// TIA Portal V20 export
// export: Created 2026-10-19T18:02:39.4342809Z, ExportSetting WithDefaults, DisplayName Totally Integrated Automation Portal, DisplayVersion V20 Update 6, DisplayName TIA Portal Openness, DisplayVersion V20 Update 6, DisplayName TIA Portal Version Control Interface, DisplayVersion V20 Update 6, DisplayName SINAMICS Startdrive Advanced, DisplayVersion V20 SP1, DisplayName SINAMICS Startdrive G130, G150, S120, S150, SINAMICS MV, G220, S200, S210, DisplayVersion V20 SP1, DisplayName SINAMICS Startdrive G110M, G120, G120C, G120D, G120P, G115D, DisplayVersion V20 SP1, DisplayName STEP 7 Professional, DisplayVersion V20 Update 6, DisplayName STEP 7 Safety, DisplayVersion V20 Update 2, DisplayName WinCC Basic/Comfort/Advanced, DisplayVersion V20 Update 6, DisplayName WinCC Unified, DisplayVersion V20 Update 6
FUNCTION "Mode_Change_F" : Void   // FC2, SCL
{ S7_Optimized_Access := 'TRUE' }
VERSION : 0.1
// stored: AutoNumber true, IsIECCheckEnabled false, SetENOAutomatically false, UDAEnableTagReadback false
   VAR_INPUT
      Mode : UInt;
   END_VAR
   VAR_TEMP
      i : UInt;
      j : UInt;
   END_VAR
BEGIN
   // REGION Change all devices
   //     "Control_DB".ECnv_Control.Instruction.Mode_Change := #Mode;
   //     "Control_DB".VTD_Control.Instruction.Mode_Change := #Mode;

   //     FOR #i := "Settings_DB".VTD_Settings.Lowest_Level TO "Settings_DB".VTD_Settings.Highest_Level DO
   //         "Control_DB".LCnv_Control.Cnv_Level_Control[#i].Cnv1_Control.Instruction.Mode_Change := #Mode;
   //         "Control_DB".LCnv_Control.Cnv_Level_Control[#i].Cnv2_Control.Instruction.Mode_Change := #Mode;
   //     END_FOR;
   // END_REGION
END_FUNCTION
